ABB RobotStudio station: Caja2Inclinada_1.rspag

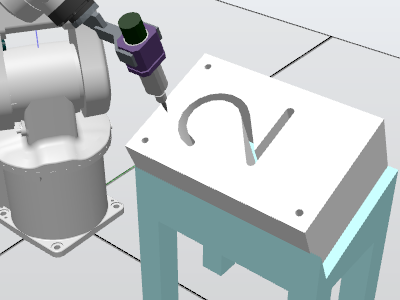
--- station ---
Station Project6 (saved by RobotStudio 26.3.11794.0)
Controller IRB120_3_58
  mechanical unit ROB_1: IRB120_3_58__01, 6 joints, base frame (0, 0, 0) mm
Layout (positions relative to the parent item):
  - IRB120_3_58__01 [mechanism, from %ABB.RobotStudio.Models.IRB120%\IRB120_3_58_G_01.rslib] at (0, 0, 0) mm; joint values [-0.5821, -0.2879, 0.4506, 0.7194, 1.0943, -0.6904] (rad or m)
  - punta [mechanism, from Components\punta.rslib] at (238.26, -106.35, 516.21) mm, rotated rx 152.86 ry 34.45 rz 164 deg
  - CajaNumero2 [part] at (585.43, -73.22, 252.41) mm, rotated rx 0 ry -22.39 rz 90.07 deg, size 188.7 x 287.5 x 103.3 mm
  - mesarRobotStudio [part] at (600, 98.92, 2.52) mm, rotated rx 0.01 ry 0 rz -179.93 deg, size 304.8 x 198.1 x 325.1 mm
Attachment: punta is attached to IRB120_3_58__01 / Link6
Collision set Conjunto de colisión_1: CajaNumero2 against punta, near miss 0 m
Targets, tools, work objects and paths stored in the station and not in the controller backup, written as RAPID:
! task T_ROB1
MODULE CalibData
  PERS tooldata MyTool:=[TRUE,[[31.792631019,0,229.638935148],[0.945518576,0,0.325568154,0]],[1,[0,0,1],[1,0,0,0],0,0,0]];
ENDMODULE


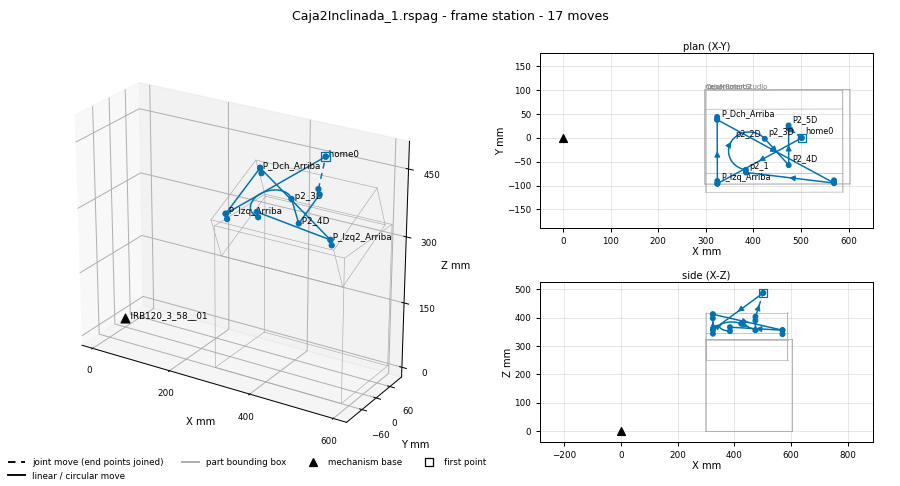
[picture p0: tool path of Caja2Inclinada_1.rspag in frame station, 17 of 17 moves have a stored position in this frame; points joined in program order, loops and branches not executed]
--- Controller Data/IRB120_3_58/RAPID/TASK1/PROGMOD/CalibData.mod ---
MODULE CalibData
    PERS tooldata punta:=[TRUE,[[24,0,172],[0.945519,0,0.325568,0]],[0.1,[0,0,1],[1,0,0,0],0,0,0]];
    TASK PERS wobjdata WOCaja:=[FALSE,TRUE,"",[[253.5,-72.5,200],[0,0.707107,0.707107,0]],[[0,0,0],[1,0,0,0]]];
    TASK PERS wobjdata cajainclinadaFernando:=[FALSE,TRUE,"",[[324.185,-94.1705,352.812],[0.137977,-0.692499,-0.695495,-0.133024]],[[0,0,0],[1,0,0,0]]];
ENDMODULE

--- Controller Data/IRB120_3_58/RAPID/TASK1/PROGMOD/Module1.mod ---
MODULE Module1
    CONST robtarget home0:=[[501.31,0,487.215],[0,0,1,0],[0,0,0,0],[9E+09,9E+09,9E+09,9E+09,9E+09,9E+09]];
    CONST robtarget P_Izq_Arriba:=[[0,0,-5],[0.707106781,-0,0,-0.707106781],[-1,0,-1,0],[9E+09,9E+09,9E+09,9E+09,9E+09,9E+09]];
    CONST robtarget P_Izq_Dentro:=[[0,0,10],[0.707106781,-0,0,-0.707106781],[-1,0,-1,0],[9E+09,9E+09,9E+09,9E+09,9E+09,9E+09]];
    CONST robtarget P_Dch_Arriba:=[[145,0,-5],[0.707106781,-0,0,-0.707106781],[0,-1,0,0],[9E+09,9E+09,9E+09,9E+09,9E+09,9E+09]];
    CONST robtarget P_Dch_Dentro:=[[145,0,10],[0.707106781,-0,0,-0.707106781],[0,-1,0,0],[9E+09,9E+09,9E+09,9E+09,9E+09,9E+09]];
    CONST robtarget P_Izq2_Arriba:=[[0,245,-5],[0.707106781,-0,0,-0.707106781],[-1,0,-1,0],[9E+09,9E+09,9E+09,9E+09,9E+09,9E+09]];
    CONST robtarget P_Izq2_Dentro:=[[0,245,10],[0.707106781,-0,0,-0.707106781],[-1,0,-1,0],[9E+09,9E+09,9E+09,9E+09,9E+09,9E+09]];
    CONST robtarget p2_1:=[[25,60,-5],[0.707106781,-0,0,-0.707106781],[-1,0,-1,0],[9E+09,9E+09,9E+09,9E+09,9E+09,9E+09]];
    CONST robtarget p2_1D:=[[25,60,10],[0.707106781,-0,0,-0.707106781],[-1,0,-1,0],[9E+09,9E+09,9E+09,9E+09,9E+09,9E+09]];
    CONST robtarget p2_2D:=[[90,30,10],[0.707106781,-0,0,-0.707106781],[0,-1,0,0],[9E+09,9E+09,9E+09,9E+09,9E+09,9E+09]];
    CONST robtarget p2_3D:=[[95,100,10],[0.707106781,-0,0,-0.707106781],[-1,0,-1,0],[9E+09,9E+09,9E+09,9E+09,9E+09,9E+09]];
    CONST robtarget P2_4D:=[[35,150,10],[0.707106781,-0,0,-0.707106781],[-1,0,-1,0],[9E+09,9E+09,9E+09,9E+09,9E+09,9E+09]];
    CONST robtarget P2_5D:=[[125,150,10],[0.707106781,-0,0,-0.707106781],[0,-1,0,0],[9E+09,9E+09,9E+09,9E+09,9E+09,9E+09]];
    CONST robtarget P2_5:=[[125,150,-5],[0.707106781,-0,0,-0.707106781],[0,-1,0,0],[9E+09,9E+09,9E+09,9E+09,9E+09,9E+09]];
    !***********************************************************
    !
    ! Module:  Module1
    !
    ! Description:
    !   <Insert description here>
    !
    ! Author: david
    !
    ! Version: 1.0
    !
    !***********************************************************


    !***********************************************************
    !
    ! Procedure main
    !
    !   This is the entry point of your program
    !
    !***********************************************************
    PROC main()
        !Add your code here
        MoveJ home0,v1000,z100,punta\WObj:=wobj0;
        MoveL P_Izq_Arriba,v200,z100,punta\WObj:=cajainclinadaFernando;
        WaitTime 2;
        MoveL P_Izq_Dentro,v20,z100,punta\WObj:=cajainclinadaFernando;
        MoveL P_Izq_Arriba,v20,z100,punta\WObj:=cajainclinadaFernando;
        MoveL P_Dch_Arriba,v20,z100,punta\WObj:=cajainclinadaFernando;
        WaitTime 2;
        MoveL P_Dch_Dentro,v20,z100,punta\WObj:=cajainclinadaFernando;
        MoveL P_Dch_Arriba,v20,z100,punta\WObj:=cajainclinadaFernando;
        MoveL P_Izq2_Arriba,v20,z100,punta\WObj:=cajainclinadaFernando;
        WaitTime 2;
        MoveL P_Izq2_Dentro,v20,z100,punta\WObj:=cajainclinadaFernando;
        MoveL P_Izq2_Arriba,v20,z100,punta\WObj:=cajainclinadaFernando;
        MoveL p2_1,v20,z100,punta\WObj:=cajainclinadaFernando;
        WaitTime 2;
        MoveL p2_1D,v10,z100,punta\WObj:=cajainclinadaFernando;
        MoveC p2_2D,p2_3D,v10,z100,punta\WObj:=cajainclinadaFernando;
        MoveL P2_4D,v10,z100,punta\WObj:=cajainclinadaFernando;
        MoveL P2_5D,v10,z100,punta\WObj:=cajainclinadaFernando;
        MoveL P2_5,v10,z100,punta\WObj:=cajainclinadaFernando;
        MoveJ home0,v20,z100,punta\WObj:=wobj0;
    ENDPROC
ENDMODULE
